# EPICS substitutions: db/Beckhoff_5XXX/ecmcEL5002.substitutions
file "ecmcEL500X-chX.template"
{
  pattern {CH_ID}
          {01   }
          {02   }
}
